(* IEC 61131-3 sources: codesys-to-s7/tests/corpus/C2S7-STD-UTIL/pos, 1 file *)

(* ---- input.st ---- *)
FUNCTION_BLOCK FB_Case
VAR
    fbBlink : BLINK;
END_VAR
fbBlink(ENABLE := TRUE);
END_FUNCTION_BLOCK
